Fanuc KAREL source: ko00079.KL

-- PROVISIONAL review KL for V770-1; original PC SHA256 132b0f544868da0e797b39d3b28c3a7e791348a7991632275557a7ac93f29669
-- Incomplete behavior may be omitted. Consult companion uncertainty JSON. Do not deploy.
PROGRAM KO00079
%NOLOCKGROUP
BEGIN
  -- UNRESOLVED_PC offsets 5-12; opcodes 9D,23
  -- UNRESOLVED_PC offsets 17-66; opcodes 27,22,1C,27,49,7E,AD,22,31,7E,4A
  -- UNRESOLVED_PC offsets 71-75; opcodes 7F
END KO00079
